TYPE E_GripperState :
(
	E_GripperState_INIT := 0,
	E_GripperState_OPENING,
	E_GripperState_OPENED,
	E_GripperState_CLOSING,
	E_GripperState_CLOSED,
	E_GripperState_UNDEFINED
);
END_TYPE

(* stored: Version 1.1.0.1, ProductVersion 3.1.4024.9
   DUT E_GripperState: Id {003cd2ae-7f7b-442c-8d6c-cea62aa79aac} *)
